# EPICS autosave request: iocs/ad/mar345-ioc/auto_settings.req
file "mar345_settings.req",       P=$(P),  R=cam1:
file "NDStdArrays_settings.req",  P=$(P),  R=image1:
file "commonPlugin_settings.req", P=$(P)
